FUNCTION_BLOCK VacuumSequence (* Composite Function Block Type *)
  (* Standard: 61499-2 *)
  (* Version 0.0, 7/2/2026, template *)
  PACKAGE Main;
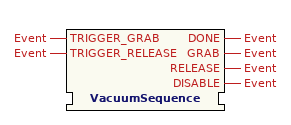
  EVENT_INPUT
    TRIGGER_GRAB;
    TRIGGER_RELEASE;
  END_EVENT
  EVENT_OUTPUT
    DONE;
    GRAB;
    RELEASE;
    DISABLE;
  END_EVENT
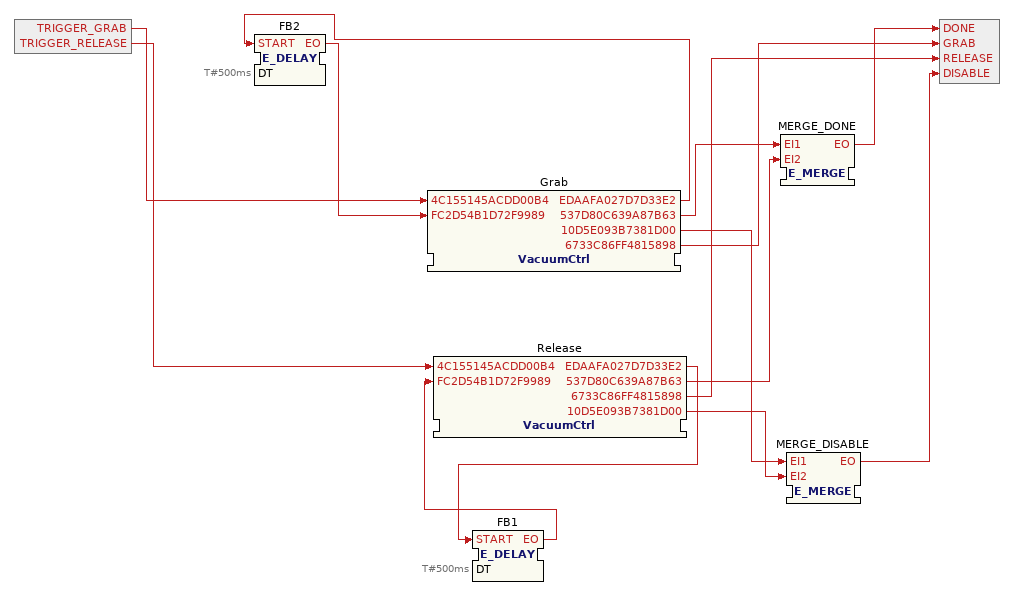
  FBS
    Grab : VacuumCtrl;
    Release : VacuumCtrl;
    MERGE_DONE : E_MERGE;
    MERGE_DISABLE : E_MERGE;
    FB1 : E_DELAY(DT := T#500ms);
    FB2 : E_DELAY(DT := T#500ms);
  END_FBS
  EVENT_CONNECTIONS
    TRIGGER_GRAB TO Grab.4C155145ACDD00B4;
    TRIGGER_RELEASE TO Release.4C155145ACDD00B4;
    FB2.EO TO Grab.FC2D54B1D72F9989;
    Grab.EDAAFA027D7D33E2 TO FB2.START;
    FB1.EO TO Release.FC2D54B1D72F9989;
    Release.EDAAFA027D7D33E2 TO FB1.START;
    Grab.537D80C639A87B63 TO MERGE_DONE.EI1;
    Release.537D80C639A87B63 TO MERGE_DONE.EI2;
    Grab.10D5E093B7381D00 TO MERGE_DISABLE.EI1;
    Grab.6733C86FF4815898 TO GRAB;
    MERGE_DONE.EO TO DONE;
    Release.6733C86FF4815898 TO RELEASE;
    MERGE_DISABLE.EO TO DISABLE;
    Release.10D5E093B7381D00 TO MERGE_DISABLE.EI2;
  END_CONNECTIONS
END_FUNCTION_BLOCK
